Fanuc KAREL source: kf00085.KL

-- PROVISIONAL review KL for V1013-1; original PC SHA256 8e0e6e1b96b2e6e6e2b08c9000e1b5beb8b6b1e2040bba08cb3abda9cd83780c
-- Incomplete behavior may be omitted. Consult companion uncertainty JSON. Do not deploy.
PROGRAM KF00085
%NOLOCKGROUP
VAR
  I : INTEGER
  J : INTEGER
  X : REAL
  Y : REAL
  B : BOOLEAN
  C : BOOLEAN
  TXT : STRING[80]
  TXT2 : STRING[80]
  STATUS : INTEGER
-- UNRESOLVED_DECL AI type=002010
-- UNRESOLVED_DECL BI type=002010
-- UNRESOLVED_DECL P type=000102
-- UNRESOLVED_DECL JP type=000199
-- UNRESOLVED_DECL PF type=000101
-- UNRESOLVED_DECL V1 type=000013
-- UNRESOLVED_DECL V2 type=000013
BEGIN
  -- UNRESOLVED_PC offsets 5-28; opcodes 49,49,AC,23
  -- UNRESOLVED_PC offsets 33-37; opcodes 7F
END KF00085
